// TIA Portal V21 export
// export: Created 2026-11-10T19:12:25.9333968Z, ExportSetting WithDefaults, DisplayName Totally Integrated Automation Portal, DisplayVersion V21 Update 3, DisplayName STEP 7 Professional, DisplayVersion V21 Update 3, DisplayName STEP 7 Safety, DisplayVersion V21, DisplayName Tech WebApplication, DisplayVersion V21, DisplayName WinCC Basic/Comfort/Advanced, DisplayVersion V21 Update 3, DisplayName WinCC Unified, DisplayVersion V21 Update 3
DATA_BLOCK "DBsTCONT_CP"   // DB33
// stored: AutoNumber true, DBAccessibleFromOPCUA true, DBAccessibleFromWebserver true, InstanceOfName TCONT_CP, OfSystemLibElement TCONT_CP, OfSystemLibVersion 1.1
TCONT_CP   // technology object, version 1.1
   // VAR_INPUT
   //    PV_IN : Real;
   //    PV_PER : Int;
   //    DISV : Real;
   //    INT_HPOS : Bool;
   //    INT_HNEG : Bool;
   //    SELECT : Int;
   // END_VAR
   // VAR_OUTPUT
   //    PV : Real;
   //    LMN : Real;
   //    LMN_PER : Int;
   //    QPULSE : Bool;
   //    QLMN_HLM : Bool;
   //    QLMN_LLM : Bool;
   //    QC_ACT : Bool;
   // END_VAR
   // VAR_IN_OUT
   //    CYCLE : Real;
   //    CYCLE_P : Real;
   //    SP_INT : Real;
   //    MAN : Real;
   //    COM_RST : Bool;
   //    MAN_ON : Bool;
   // END_VAR
   // VAR RETAIN
   //    DEADB_W : Real;
   //    I_ITLVAL : Real;
   //    LMN_HLM : Real;
   //    LMN_LLM : Real;
   //    PV_FAC : Real;
   //    PV_OFFS : Real;
   //    LMN_FAC : Real;
   //    LMN_OFFS : Real;
   //    PER_TM : Real;
   //    P_B_TM : Real;
   //    TUN_DLMN : Real;
   //    PER_MODE : Int;
   //    PVPER_ON : Bool;
   //    I_ITL_ON : Bool;
   //    PULSE_ON : Bool;
   //    TUN_KEEP : Bool;
   //    ER : Real;
   //    LMN_P : Real;
   //    LMN_I : Real;
   //    LMN_D : Real;
   //    PHASE : Int;
   //    STATUS_H : Int;
   //    STATUS_D : Int;
   //    QTUN_RUN : Bool;
   //    PI_CON { S7_SetPoint := 'True'} : TCONTCP_PI_CON;
   //    PID_CON { S7_SetPoint := 'True'} : TCONTCP_PID_CON;
   //    PAR_SAVE { S7_SetPoint := 'True'} : TCONTCP_PAR_SAVE;
   //    PFAC_SP : Real;
   //    GAIN : Real;
   //    TI : Real;
   //    TD : Real;
   //    D_F : Real;
   //    CON_ZONE : Real;
   //    CONZ_ON : Bool;
   //    TUN_ON : Bool;
   //    TUN_ST : Bool;
   //    UNDO_PAR : Bool;
   //    SAVE_PAR : Bool;
   //    LOAD_PID : Bool;
   //    PID_ON : Bool;
   //    GAIN_P : Real;
   //    TU : Real;
   //    TA : Real;
   //    KIG : Real;
   //    N_PTN : Real;
   //    TM_LAG_P : Real;
   //    T_P_INF : Real;
   //    P_INF : Real;
   //    LMN0 : Real;
   //    PV0 : Real;
   //    PVDT0 : Real;
   //    PVDT : Real;
   //    PVDT_MAX : Real;
   //    NOI_PVDT : Real;
   //    NOISE_PV : Real;
   //    FIL_CYC : Int;
   //    POI_CMAX : Int;
   //    POI_CYCL : Int;
   //    sctFil : Int;
   //    srPv : Real;
   //    srNoise : Real;
   //    srPvdt2 : Real;
   //    srPvdtMax2 : Real;
   //    srNoise2 : Real;
   //    srPvOld2 : Real;
   //    siStatus : Int;
   //    siSpDir : Int;
   //    srTime : Real;
   //    sPvOld : Real;
   //    sSpOld : Real;
   //    srPvMin : Real;
   //    srPVsim : Real;
   //    srEffDlmn : Real;
   //    sInvAlt : Real;
   //    sIanteilAlt : Real;
   //    sRestInt : Real;
   //    sRestDif : Real;
   //    sRueck : Real;
   //    sLmn : Real;
   //    spassPTm : Real;
   //    sCycTmPass : Real;
   //    sPTm : Real;
   //    srOptLmn : Real;
   //    sbOptLmn : Bool;
   //    sbConzOn : Bool;
   //    sbSpChange : Bool;
   //    sbReOpt : Bool;
   //    sLmnHlmOld : Real;
   //    sLmnLlmOld : Real;
   //    srDiffSp : Real;
   //    siTime : DInt;
   //    siCycle : DInt;
   //    siCycleP : DInt;
   //    siPulsFil : Int;
   //    srPulsPv : Real;
   //    srDPvdt : Real;
   //    srDPvdt2 : Real;
   //    sNpInf : Real;
   //    sCycleM : Real;
   //    sGf11_30 : Real;
   //    sGf12_30 : Real;
   //    sGf21_30 : Real;
   //    sGf22_30 : Real;
   //    sPv0Sim_30 : Real;
   //    srPVsim3_30 : Real;
   //    srPVsim2_30 : Real;
   //    srPVsim1_30 : Real;
   //    srDelPvsim_30 : Real;
   //    sGf11_20 : Real;
   //    sGf12_20 : Real;
   //    sGf21_20 : Real;
   //    sGf22_20 : Real;
   //    sPv0Sim_20 : Real;
   //    srPVsim2_20 : Real;
   //    srPVsim1_20 : Real;
   //    srDelPvsim_20 : Real;
   //    sGf11_15 : Real;
   //    sGf12_15 : Real;
   //    sGf21_15 : Real;
   //    sGf22_15 : Real;
   //    sPv0Sim_15 : Real;
   //    srPVsim2_15 : Real;
   //    srPVsim1_15 : Real;
   //    srDelPvsim_15 : Real;
   // END_VAR
BEGIN
END_DATA_BLOCK
